(* IEC 61131-3 sources: llm-plc-st-eval/data/definitivo/claude-sonnet-4-6/A2/zero_shot, 3 files *)

(* ---- ejec_1.st ---- *)
```pascal
FUNCTION_BLOCK FB_Batch

VAR_INPUT
    nivelA    : BOOL;   (* Sensor nivel componente A alcanzado *)
    nivelB    : BOOL;   (* Sensor nivel componente B alcanzado *)
    nivelVacio : BOOL;  (* Sensor reactor vacío *)
    btnInicio : BOOL;   (* Botón inicio receta (flanco no requerido, nivel) *)
    btnAbort  : BOOL;   (* Botón abort *)
    temp      : REAL;   (* Temperatura actual del reactor *)
END_VAR

VAR_OUTPUT
    vA        : BOOL;   (* Válvula componente A *)
    vB        : BOOL;   (* Válvula componente B *)
    calentador : BOOL;  (* Calentador *)
    mezclador : BOOL;   (* Mezclador *)
    vDescarga : BOOL;   (* Válvula de descarga *)
    fase      : INT;    (* Fase activa: 0=reposo, 1-5=fases receta *)
END_VAR

VAR
    timerMezcla   : TON;        (* Temporizador fase 4 mezcla *)
    abortActivo   : BOOL;       (* Indica que se está ejecutando un abort *)
    btnInicioAnterior : BOOL;   (* Flanco ascendente btnInicio *)
    btnAbortAnterior  : BOOL;   (* Flanco ascendente btnAbort *)
    flancoInicio  : BOOL;       (* Flanco detectado btnInicio *)
    flancoAbort   : BOOL;       (* Flanco detectado btnAbort *)
END_VAR

(* ─── Detección de flancos ascendentes ─────────────────────────────────── *)
flancoInicio := btnInicio AND NOT btnInicioAnterior;
flancoAbort  := btnAbort  AND NOT btnAbortAnterior;

(* ─── Lógica principal por fase ─────────────────────────────────────────── *)

(* --- Gestión de ABORT (fases 1 a 5) ------------------------------------ *)
IF flancoAbort AND (fase >= 1) AND (fase <= 5) THEN
    abortActivo := TRUE;

    (* Apagar actuadores de proceso inmediatamente *)
    vA         := FALSE;
    vB         := FALSE;
    calentador := FALSE;
    mezclador  := FALSE;

    (* Decidir siguiente estado *)
    IF fase = 5 THEN
        (* Ya estamos descargando: continuar fase 5 sin cambio *)
        (* abortActivo queda TRUE para que al vaciar vuelva a reposo *)
        (* No se cambia fase *)
    ELSIF nivelVacio THEN
        (* Reactor ya vacío: ir directamente a reposo *)
        vDescarga  := FALSE;
        fase       := 0;
        abortActivo := FALSE;
    ELSE
        (* Hay producto: ir a fase 5 para descargar *)
        fase := 5;
    END_IF;
END_IF;

(* --- Máquina de estados ------------------------------------------------- *)
CASE fase OF

    (* ── FASE 0: Reposo ─────────────────────────────────────────────── *)
    0:
        (* Asegurar todas las salidas apagadas *)
        vA         := FALSE;
        vB         := FALSE;
        calentador := FALSE;
        mezclador  := FALSE;
        vDescarga  := FALSE;
        abortActivo := FALSE;

        (* Arranque solo con flanco de btnInicio *)
        IF flancoInicio THEN
            fase := 1;
        END_IF;

    (* ── FASE 1: Dosificar componente A ─────────────────────────────── *)
    1:
        vA := TRUE;

        IF nivelA THEN
            vA   := FALSE;
            fase := 2;
        END_IF;

    (* ── FASE 2: Dosificar componente B ─────────────────────────────── *)
    2:
        vB := TRUE;

        IF nivelB THEN
            vB   := FALSE;
            fase := 3;
        END_IF;

    (* ── FASE 3: Calentar hasta 60 °C ───────────────────────────────── *)
    3:
        calentador := TRUE;

        IF temp >= 60.0 THEN
            calentador := FALSE;
            fase       := 4;
            (* Reiniciar temporizador antes de entrar en fase 4 *)
            timerMezcla(IN := FALSE, PT := T#120S);
        END_IF;

    (* ── FASE 4: Mezclar 120 segundos ───────────────────────────────── *)
    4:
        mezclador := TRUE;
        timerMezcla(IN := TRUE, PT := T#120S);

        IF timerMezcla.Q THEN
            mezclador := FALSE;
            timerMezcla(IN := FALSE, PT := T#120S); (* Reset timer *)
            fase := 5;
        END_IF;

    (* ── FASE 5: Descargar hasta reactor vacío ──────────────────────── *)
    5:
        vDescarga := TRUE;

        IF nivelVacio THEN
            vDescarga   := FALSE;
            fase        := 0;
            abortActivo := FALSE;
        END_IF;

    (* ── Estado no definido: volver a reposo ────────────────────────── *)
    ELSE:
        fase := 0;

END_CASE;

(* ─── Actualizar memoria de flancos ─────────────────────────────────────── *)
btnInicioAnterior := btnInicio;
btnAbortAnterior  := btnAbort;
```

(* ---- ejec_2.st ---- *)
```pascal
FUNCTION_BLOCK FB_Batch
VAR_INPUT
    nivelA    : BOOL;   (* Sensor nivel componente A alcanzado *)
    nivelB    : BOOL;   (* Sensor nivel componente B alcanzado *)
    nivelVacio: BOOL;   (* Sensor reactor vacío *)
    btnInicio : BOOL;   (* Botón inicio receta (flanco no requerido, nivel) *)
    btnAbort  : BOOL;   (* Botón abort *)
    temp      : REAL;   (* Temperatura actual del reactor *)
END_VAR

VAR_OUTPUT
    vA        : BOOL;   (* Válvula componente A *)
    vB        : BOOL;   (* Válvula componente B *)
    calentador: BOOL;   (* Calentador *)
    mezclador : BOOL;   (* Mezclador *)
    vDescarga : BOOL;   (* Válvula de descarga *)
    fase      : INT;    (* Fase activa: 0=reposo, 1-5=fases receta *)
END_VAR

VAR
    timerMezcla   : TON;            (* Temporizador fase 4 mezcla *)
    abortando     : BOOL;           (* Indica que se está ejecutando un abort *)
    btnInicio_prev: BOOL;           (* Valor anterior de btnInicio para flanco *)
    btnAbort_prev : BOOL;           (* Valor anterior de btnAbort para flanco *)
    btnInicio_re  : BOOL;           (* Flanco ascendente btnInicio *)
    btnAbort_re   : BOOL;           (* Flanco ascendente btnAbort *)
END_VAR

(* ─────────────────────────────────────────────
   Detección de flancos ascendentes
   ───────────────────────────────────────────── *)
btnInicio_re := btnInicio AND NOT btnInicio_prev;
btnAbort_re  := btnAbort  AND NOT btnAbort_prev;

(* ─────────────────────────────────────────────
   Lógica principal de fases
   ───────────────────────────────────────────── *)
CASE fase OF

    (* ── FASE 0: Reposo ── *)
    0:
        abortando := FALSE;

        (* Arranque solo desde reposo, con flanco de btnInicio *)
        IF btnInicio_re THEN
            fase := 1;
        END_IF;
        (* btnAbort en reposo no tiene efecto *)

    (* ── FASE 1: Dosificar componente A ── *)
    1:
        IF btnAbort_re THEN
            abortando := TRUE;
            (* Cerrar actuadores inmediatamente *)
            vA        := FALSE;
            vB        := FALSE;
            calentador:= FALSE;
            mezclador := FALSE;
            (* Decidir si hay que descargar *)
            IF NOT nivelVacio THEN
                fase := 5;  (* Hay producto: descargar *)
            ELSE
                fase := 0;  (* Reactor ya vacío: reposo *)
            END_IF;
        ELSIF nivelA THEN
            fase := 2;      (* Nivel A alcanzado: siguiente fase *)
        END_IF;

    (* ── FASE 2: Dosificar componente B ── *)
    2:
        IF btnAbort_re THEN
            abortando := TRUE;
            vA        := FALSE;
            vB        := FALSE;
            calentador:= FALSE;
            mezclador := FALSE;
            IF NOT nivelVacio THEN
                fase := 5;
            ELSE
                fase := 0;
            END_IF;
        ELSIF nivelB THEN
            fase := 3;      (* Nivel B alcanzado: siguiente fase *)
        END_IF;

    (* ── FASE 3: Calentar ── *)
    3:
        IF btnAbort_re THEN
            abortando := TRUE;
            vA        := FALSE;
            vB        := FALSE;
            calentador:= FALSE;
            mezclador := FALSE;
            IF NOT nivelVacio THEN
                fase := 5;
            ELSE
                fase := 0;
            END_IF;
        ELSIF temp >= 60.0 THEN
            fase := 4;      (* Temperatura alcanzada: siguiente fase *)
        END_IF;

    (* ── FASE 4: Mezclar 120 s ── *)
    4:
        IF btnAbort_re THEN
            abortando := TRUE;
            vA        := FALSE;
            vB        := FALSE;
            calentador:= FALSE;
            mezclador := FALSE;
            timerMezcla(IN := FALSE);  (* Resetear temporizador *)
            IF NOT nivelVacio THEN
                fase := 5;
            ELSE
                fase := 0;
            END_IF;
        ELSIF timerMezcla.Q THEN
            timerMezcla(IN := FALSE);  (* Resetear temporizador *)
            fase := 5;                 (* Tiempo cumplido: descargar *)
        END_IF;

    (* ── FASE 5: Descargar ── *)
    5:
        (* Un abort durante la descarga continúa la descarga;
           solo se marca abortando si aún no estaba activo *)
        IF btnAbort_re AND NOT abortando THEN
            abortando := TRUE;
            (* Los demás actuadores ya deben estar apagados,
               pero se asegura por si el abort ocurre en fase 5 normal *)
            vA        := FALSE;
            vB        := FALSE;
            calentador:= FALSE;
            mezclador := FALSE;
        END_IF;

        IF nivelVacio THEN
            fase := 0;      (* Reactor vacío: volver a reposo *)
        END_IF;

END_CASE;

(* ─────────────────────────────────────────────
   Asignación de salidas según fase activa
   ───────────────────────────────────────────── *)
CASE fase OF
    0:  (* Reposo: todo apagado *)
        vA         := FALSE;
        vB         := FALSE;
        calentador := FALSE;
        mezclador  := FALSE;
        vDescarga  := FALSE;
        timerMezcla(IN := FALSE);

    1:  (* Dosificar A *)
        vA         := TRUE;
        vB         := FALSE;
        calentador := FALSE;
        mezclador  := FALSE;
        vDescarga  := FALSE;
        timerMezcla(IN := FALSE);

    2:  (* Dosificar B *)
        vA         := FALSE;
        vB         := TRUE;
        calentador := FALSE;
        mezclador  := FALSE;
        vDescarga  := FALSE;
        timerMezcla(IN := FALSE);

    3:  (* Calentar *)
        vA         := FALSE;
        vB         := FALSE;
        calentador := TRUE;
        mezclador  := FALSE;
        vDescarga  := FALSE;
        timerMezcla(IN := FALSE);

    4:  (* Mezclar *)
        vA         := FALSE;
        vB         := FALSE;
        calentador := FALSE;
        mezclador  := TRUE;
        vDescarga  := FALSE;
        timerMezcla(IN := TRUE, PT := T#120S);  (* Activar temporizador *)

    5:  (* Descargar *)
        vA         := FALSE;
        vB         := FALSE;
        calentador := FALSE;
        mezclador  := FALSE;
        vDescarga  := TRUE;
        timerMezcla(IN := FALSE);

END_CASE;

(* ─────────────────────────────────────────────
   Actualizar valores previos para próximo ciclo
   ───────────────────────────────────────────── *)
btnInicio_prev := btnInicio;
btnAbort_prev  := btnAbort;
```

(* ---- ejec_3.st ---- *)
```pascal
FUNCTION_BLOCK FB_Batch

VAR_INPUT
    nivelA    : BOOL;   (* Sensor nivel componente A alcanzado *)
    nivelB    : BOOL;   (* Sensor nivel componente B alcanzado *)
    nivelVacio: BOOL;   (* Sensor reactor vacío *)
    btnInicio : BOOL;   (* Botón inicio receta (flanco no requerido, nivel) *)
    btnAbort  : BOOL;   (* Botón abort *)
    temp      : REAL;   (* Temperatura actual del reactor *)
END_VAR

VAR_OUTPUT
    vA        : BOOL;   (* Válvula componente A *)
    vB        : BOOL;   (* Válvula componente B *)
    calentador: BOOL;   (* Calentador *)
    mezclador : BOOL;   (* Mezclador *)
    vDescarga : BOOL;   (* Válvula de descarga *)
    fase      : INT;    (* Fase activa: 0=reposo, 1-5=receta *)
END_VAR

VAR
    timerMezcla   : TON;        (* Temporizador fase 4 mezcla *)
    abortando     : BOOL;       (* Indica que se está ejecutando un abort *)
    btnInicioAnterior : BOOL;   (* Para detección de flanco ascendente btnInicio *)
    btnAbortAnterior  : BOOL;   (* Para detección de flanco ascendente btnAbort *)
    flancoInicio  : BOOL;       (* Flanco ascendente btnInicio *)
    flancoAbort   : BOOL;       (* Flanco ascendente btnAbort *)
END_VAR

(* ─────────────────────────────────────────────
   Detección de flancos ascendentes
   ───────────────────────────────────────────── *)
flancoInicio := btnInicio AND NOT btnInicioAnterior;
flancoAbort  := btnAbort  AND NOT btnAbortAnterior;

(* ─────────────────────────────────────────────
   Lógica principal por fases
   ───────────────────────────────────────────── *)
CASE fase OF

    (* ── FASE 0: Reposo ── *)
    0:
        abortando := FALSE;

        (* Arranque solo desde reposo, con flanco *)
        IF flancoInicio THEN
            fase := 1;
        END_IF;
        (* btnAbort en reposo no tiene efecto *)

    (* ── FASE 1: Dosificar componente A ── *)
    1:
        IF flancoAbort THEN
            (* Abort: cerrar actuadores y decidir si descargar *)
            abortando := TRUE;
            IF NOT nivelVacio THEN
                fase := 5;      (* Hay producto → descargar *)
            ELSE
                fase := 0;      (* Reactor ya vacío → reposo *)
            END_IF;
        ELSIF nivelA THEN
            fase := 2;          (* Nivel A alcanzado → siguiente fase *)
        END_IF;

    (* ── FASE 2: Dosificar componente B ── *)
    2:
        IF flancoAbort THEN
            abortando := TRUE;
            IF NOT nivelVacio THEN
                fase := 5;
            ELSE
                fase := 0;
            END_IF;
        ELSIF nivelB THEN
            fase := 3;          (* Nivel B alcanzado → siguiente fase *)
        END_IF;

    (* ── FASE 3: Calentar hasta 60 °C ── *)
    3:
        IF flancoAbort THEN
            abortando := TRUE;
            IF NOT nivelVacio THEN
                fase := 5;
            ELSE
                fase := 0;
            END_IF;
        ELSIF temp >= 60.0 THEN
            fase := 4;          (* Temperatura alcanzada → siguiente fase *)
        END_IF;

    (* ── FASE 4: Mezclar 120 segundos ── *)
    4:
        IF flancoAbort THEN
            abortando := TRUE;
            timerMezcla(IN := FALSE);   (* Resetear temporizador *)
            IF NOT nivelVacio THEN
                fase := 5;
            ELSE
                fase := 0;
            END_IF;
        ELSIF timerMezcla.Q THEN
            timerMezcla(IN := FALSE);   (* Resetear temporizador *)
            fase := 5;                  (* Tiempo cumplido → descargar *)
        END_IF;

    (* ── FASE 5: Descargar ── *)
    5:
        (* Un abort durante fase 5 continúa la descarga normalmente *)
        (* Solo se marca abortando si vino de otra fase; aquí no se interrumpe *)
        IF nivelVacio THEN
            fase := 0;          (* Reactor vacío → reposo *)
            abortando := FALSE;
        END_IF;
        (* flancoAbort en fase 5 se ignora (descarga continúa) *)

END_CASE;

(* ─────────────────────────────────────────────
   Asignación de salidas según fase activa
   ───────────────────────────────────────────── *)

(* Válvula A: abierta solo en fase 1 normal (no en abort) *)
vA := (fase = 1) AND NOT abortando;

(* Válvula B: abierta solo en fase 2 normal *)
vB := (fase = 2) AND NOT abortando;

(* Calentador: activo solo en fase 3 normal *)
calentador := (fase = 3) AND NOT abortando;

(* Mezclador: activo solo en fase 4 normal *)
mezclador := (fase = 4) AND NOT abortando;

(* Válvula descarga: abierta en fase 5 (normal o por abort) *)
vDescarga := (fase = 5);

(* ─────────────────────────────────────────────
   Temporizador mezcla (fase 4)
   ───────────────────────────────────────────── *)
timerMezcla(IN := (fase = 4) AND NOT abortando, PT := T#120S);

(* ─────────────────────────────────────────────
   Actualizar estados anteriores de botones
   ───────────────────────────────────────────── *)
btnInicioAnterior := btnInicio;
btnAbortAnterior  := btnAbort;

END_FUNCTION_BLOCK
```
